// TIA Portal V20 program export: 0 tag tables, 0 data types, 0 data blocks, 1 code blocks (in call order from the OBs), 0 instance data blocks

ORGANIZATION_BLOCK "Main"   // OB1, LAD, ProgramCycle
TITLE = "Main Program Sweep (Cycle)"
{ S7_Optimized_Access := 'TRUE' }
// stored: SetENOAutomatically false
   VAR_INPUT
      Initial_Call : Bool;
      Remanence : Bool;
   END_VAR
BEGIN

REGION Network 1
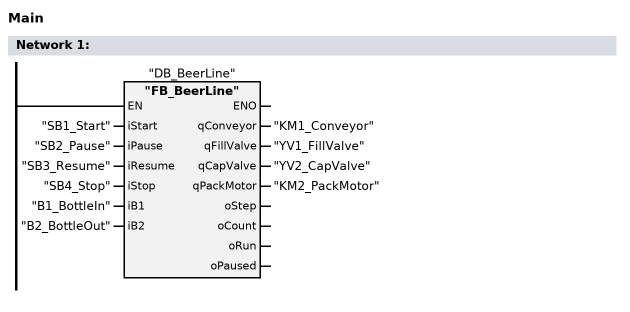
   RUNG wire#powerrail
      "DB_BeerLine"(iStart := "SB1_Start", iPause := "SB2_Pause", iResume := "SB3_Resume", iStop := "SB4_Stop", iB1 := "B1_BottleIn", iB2 := "B2_BottleOut", qConveyor => "KM1_Conveyor", qFillValve => "YV1_FillValve", qCapValve => "YV2_CapValve", qPackMotor => "KM2_PackMotor", oStep =>, oCount =>, oRun =>, oPaused =>)
   END_RUNG
   // the same network as SCL:
   "DB_BeerLine"(iStart := "SB1_Start",   // "FB_BeerLine"
                 iPause := "SB2_Pause",
                 iResume := "SB3_Resume",
                 iStop := "SB4_Stop",
                 iB1 := "B1_BottleIn",
                 iB2 := "B2_BottleOut",
                 qConveyor => "KM1_Conveyor",
                 qFillValve => "YV1_FillValve",
                 qCapValve => "YV2_CapValve",
                 qPackMotor => "KM2_PackMotor");
END_REGION
END_ORGANIZATION_BLOCK
